// TIA Portal V21 export
DATA_BLOCK "DB_Recipes"   // DB3
TITLE = Rezeptspeicher / Recipe storage
// Array-DB mit zehn Abfüllrezepten / Array DB holding ten filling recipes
   STRUCT
      DB_Recipes : Array[0..9] of "UDT_Recipe";
   END_STRUCT;
BEGIN
END_DATA_BLOCK
